// TIA Portal V21 export
TextList "TL_State"  ListRange=Decimal
  TextListEntry   Text="OFF"
  TextListEntry   From=1, To=1, Text="INIT"
